FUNCTION_BLOCK Controle_Necessidade (* Necessidade de equipamentos por faixas de nivel (padrao Necessidade_2_Equipamentos do legado) *)
  (* Standard: 61499-2 *)
  (* Version 1.0, 21/10/2026, Hidryco, Hidryco, 1.0: Necessidade de equipamentos por faixas de nivel (padrao Necessidade_2_Equipamentos do legado) *)
  PACKAGE Hidryco.HidrycoLib;
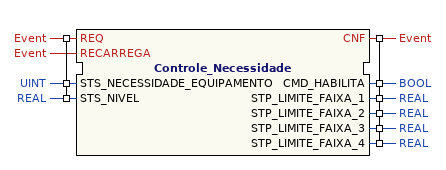
  EVENT_INPUT
    REQ WITH STS_NECESSIDADE_EQUIPAMENTO, STS_NIVEL; (* Status vindo do processo *)
    RECARREGA; (* Reenvia os ajustes persistentes (chamado no fim do INIT do processo) *)
  END_EVENT
  EVENT_OUTPUT
    CNF WITH CMD_HABILITA, STP_LIMITE_FAIXA_1, STP_LIMITE_FAIXA_2, STP_LIMITE_FAIXA_3, STP_LIMITE_FAIXA_4; (* Ajustes para o processo (mudanca na IHM, OPC UA ou recarga) *)
  END_EVENT
  VAR_INPUT
    STS_NECESSIDADE_EQUIPAMENTO : UINT; (* Equipamentos pedidos pelas faixas *)
    STS_NIVEL : REAL; (* Nivel comparado com as faixas (% da altura) *)
  END_VAR
  VAR_OUTPUT
    CMD_HABILITA : BOOL; (* Habilitado *)
    STP_LIMITE_FAIXA_1 : REAL; (* Limite da faixa 1 *)
    STP_LIMITE_FAIXA_2 : REAL; (* Limite da faixa 2 *)
    STP_LIMITE_FAIXA_3 : REAL; (* Limite da faixa 3 *)
    STP_LIMITE_FAIXA_4 : REAL; (* Limite da faixa 4 *)
  END_VAR
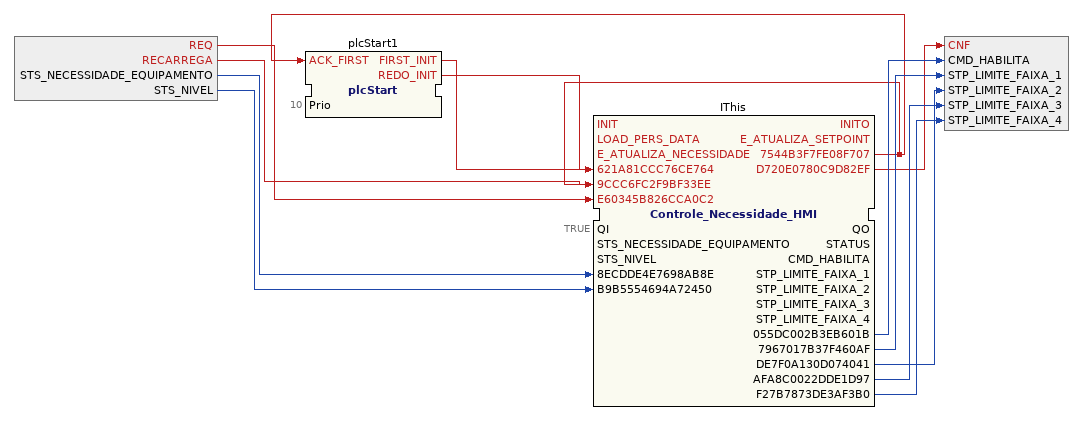
  FBS
    IThis : Controle_Necessidade_HMI(QI := TRUE);
    plcStart1 : plcStart(Prio := 10);
  END_FBS
  EVENT_CONNECTIONS
    plcStart1.FIRST_INIT TO IThis.621A81CCC76CE764;
    plcStart1.REDO_INIT TO IThis.621A81CCC76CE764;
    IThis.7544B3F7FE08F707 TO IThis.9CCC6FC2F9BF33EE;
    IThis.7544B3F7FE08F707 TO plcStart1.ACK_FIRST;
    RECARREGA TO IThis.9CCC6FC2F9BF33EE;
    IThis.D720E0780C9D82EF TO CNF;
    REQ TO IThis.E60345B826CCA0C2;
  END_CONNECTIONS
  DATA_CONNECTIONS
    IThis.055DC002B3EB601B TO CMD_HABILITA;
    IThis.7967017B37F460AF TO STP_LIMITE_FAIXA_1;
    IThis.DE7F0A130D074041 TO STP_LIMITE_FAIXA_2;
    IThis.AFA8C0022DDE1D97 TO STP_LIMITE_FAIXA_3;
    IThis.F27B7873DE3AF3B0 TO STP_LIMITE_FAIXA_4;
    STS_NECESSIDADE_EQUIPAMENTO TO IThis.8ECDDE4E7698AB8E;
    STS_NIVEL TO IThis.B9B5554694A72450;
  END_CONNECTIONS
END_FUNCTION_BLOCK
